ADAPTER AContract (* An adapter: one connection from a primitive's contract (SC_, the plug) to its run (SKILL_Run, the socket) that carries what the contract says: at the start what to do and whether it may start, at each new state of the equipment whether it is done and may go on. Technical: What a skill primitive's contract (SC_, the plug) tells its run (SKILL_Run, the socket): at START what to do and whether it may start, at SAMPLE whether the newest state of the equipment ends the run *)
  (* Standard: 61499-2 *)
  (* Version 0.1, 2026-09-28, Project contributors, AAU Smart Production Lab *)
  PACKAGE modlib;
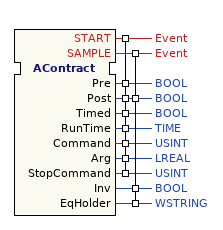
  EVENT_OUTPUT
    START WITH Pre, Post, Timed, RunTime, Command, Arg, StopCommand; (* A run starts: what to do (Command, Arg, RunTime, StopCommand) and whether it may (Pre) *)
    SAMPLE WITH Post, Inv, EqHolder; (* The equipment's newest state, judged: is the skill done (Post), may it go on (Inv) *)
  END_EVENT
  VAR_OUTPUT
    Pre : BOOL;
    Post : BOOL;
    Timed : BOOL;
    RunTime : TIME;
    Command : USINT;
    Arg : LREAL;
    StopCommand : USINT;
    Inv : BOOL;
    EqHolder : WSTRING; (* Who holds the equipment now (empty: free) *)
  END_VAR
END_ADAPTER
